(* IEC 61131-3 sources: st-fmt/tests/fixtures/realworld, 8 files *)

(* ---- analog_input_udt.expected.st ---- *)
TYPE
analog_input_8channel_udt : STRUCT
    {attribute 'symbol' := 'read'}
    position1       : REAL;
    {attribute 'symbol' := 'read'}
    position1_fault : BOOL;
    {attribute 'symbol' := 'read'}
    position2       : REAL;
    {attribute 'symbol' := 'read'}
    position2_fault : BOOL;
    {attribute 'symbol' := 'read'}
    position3       : REAL;
    {attribute 'symbol' := 'read'}
    position3_fault : BOOL;
    {attribute 'symbol' := 'read'}
    position4       : REAL;
    {attribute 'symbol' := 'read'}
    position4_fault : BOOL;
    {attribute 'symbol' := 'read'}
    position5       : REAL;
    {attribute 'symbol' := 'read'}
    position5_fault : BOOL;
    {attribute 'symbol' := 'read'}
    position6       : REAL;
    {attribute 'symbol' := 'read'}
    position6_fault : BOOL;
    {attribute 'symbol' := 'read'}
    position7       : REAL;
    {attribute 'symbol' := 'read'}
    position7_fault : BOOL;
    {attribute 'symbol' := 'read'}
    position8       : REAL;
    {attribute 'symbol' := 'read'}
    position8_fault : BOOL;
END_STRUCT
END_TYPE

(* ---- analog_input_udt.st ---- *)
TYPE analog_input_8channel_udt :
STRUCT
	{attribute 'symbol' := 'read'}
	position1: REAL;
	{attribute 'symbol' := 'read'}
	position1_fault: BOOL;
	{attribute 'symbol' := 'read'}
	position2: REAL;
	{attribute 'symbol' := 'read'}
	position2_fault: BOOL;
	{attribute 'symbol' := 'read'}
	position3: REAL;
	{attribute 'symbol' := 'read'}
	position3_fault: BOOL;
	{attribute 'symbol' := 'read'}
	position4: REAL;
	{attribute 'symbol' := 'read'}
	position4_fault: BOOL;
	{attribute 'symbol' := 'read'}
	position5: REAL;
	{attribute 'symbol' := 'read'}
	position5_fault: BOOL;
	{attribute 'symbol' := 'read'}
	position6: REAL;
	{attribute 'symbol' := 'read'}
	position6_fault: BOOL;
	{attribute 'symbol' := 'read'}
	position7: REAL;
	{attribute 'symbol' := 'read'}
	position7_fault: BOOL;
	{attribute 'symbol' := 'read'}
	position8: REAL;
	{attribute 'symbol' := 'read'}
	position8_fault: BOOL;
END_STRUCT
END_TYPE

(* ---- test_error_message.expected.st ---- *)
{attribute 'pack_mode':='1'}
TYPE
TestErrorMessage : STRUCT
    step    : INT;
    message : STRING[512];
END_STRUCT
END_TYPE

(* ---- test_error_message.st ---- *)
{attribute 'pack_mode':='1'}
TYPE TestErrorMessage :
STRUCT
	step: INT;
	message: STRING[512];
END_STRUCT
END_TYPE

(* ---- debounce.expected.st ---- *)
FUNCTION_BLOCK debounce
VAR_INPUT
    input         : BOOL;
    debounce_time : TIME;
END_VAR
VAR_OUTPUT
    output : BOOL;
END_VAR
VAR
    _debounce_timer : TON;
END_VAR

_debounce_timer(in := input XOR output, PT := debounce_time);
IF _debounce_timer.Q THEN
    output := input;
ELSE
    output := output;
END_IF

END_FUNCTION_BLOCK

(* ---- debounce.st ---- *)
FUNCTION_BLOCK debounce
VAR_INPUT
	input: BOOL;
	debounce_time: TIME;
END_VAR
VAR_OUTPUT
	output: BOOL;
END_VAR
VAR
	_debounce_timer: TON;
END_VAR

_debounce_timer(in := input XOR output, PT := debounce_time);
IF _debounce_timer.Q THEN
	output := input;
ELSE
	output := output;
END_IF;
END_FUNCTION_BLOCK

(* ---- base_test_run.expected.st ---- *)
METHOD Run : BOOL
VAR_INPUT
    duration : TIME := T#0s;
END_VAR
VAR_OUTPUT
    pos : INT;
END_VAR

(*
	Checks the active step and returns true if active.
	Sets the delay if active.
	Calculates the amount of steps in the test.
	Calculates the total amount of delay time for the test.
*)
IF NOT _inizialized THEN
    _error := TRUE;
    SetMessage('Run method called without initialization. Init method needs to be called first.');
END_IF

Run            := CurrentStep = _scan_index AND State = TestState.Running;
OnEntry        := Run AND _step_previous = CurrentStep;
_step_previous := CurrentStep;
pos            := _scan_index;
IF Run THEN
    _delay := duration;
END_IF

_scan_index := _scan_index + 1;
IF State = TestState.Starting AND _scan_index > TotalStepCount THEN
    TotalStepCount := _scan_index;
    IF _loop_index = 0 THEN
        TestDurationExpected := TestDurationExpected + MAX(duration, TO_TIME(_cycle_time));
    ELSE
        _loop_time[_loop_index] := _loop_time[_loop_index] + MAX(duration, TO_TIME(_cycle_time));
    END_IF
END_IF

(* ---- base_test_run.st ---- *)
METHOD Run : BOOL
VAR_INPUT
	duration : TIME := T#0s;
END_VAR
VAR_OUTPUT
	pos: INT;
END_VAR

(*
	Checks the active step and returns true if active.
	Sets the delay if active.
	Calculates the amount of steps in the test.
	Calculates the total amount of delay time for the test.
*)
IF NOT _inizialized THEN
	_error := TRUE;
	SetMessage('Run method called without initialization. Init method needs to be called first.');
END_IF;

Run := CurrentStep = _scan_index AND State = TestState.Running;
OnEntry := Run AND _step_previous = CurrentStep;
_step_previous := CurrentStep;
pos := _scan_index;
IF Run THEN
	_delay := duration;
END_IF;
_scan_index := _scan_index + 1;
IF State = TestState.Starting AND  _scan_index > TotalStepCount THEN
	TotalStepCount := _scan_index;
	IF _loop_index = 0 THEN
		TestDurationExpected := TestDurationExpected + MAX(duration, TO_TIME(_cycle_time));
	ELSE
		_loop_time[_loop_index] := _loop_time[_loop_index] + MAX(duration, TO_TIME(_cycle_time));
	END_IF;
END_IF;
